INTERFACE I_Cyclic EXTENDS __SYSTEM.IQueryInterface

// Called once per scan, by whoever owns this block's place in the call order.

METHOD CyclicLogic
END_METHOD

END_INTERFACE

(* stored: Version 1.1.0.1
   Itf I_Cyclic: Id {fb9a048c-fd1e-40db-a4c6-d3970535ecf2}
   Method CyclicLogic: Id {91ff5771-17cc-4645-ac61-cbceda3c18ac} *)
